// TIA Portal project "latest plc" (V21)

(* hardware
DEVICE "S7-1200 station_1"  S7-1200 Station
   slot 0: "Rack_0"  S7-1200 Rack  Rack  V1.0
   slot 1: "PLC_1"  CPU 1214C DC/DC/DC  6ES7 214-1AG40-0XB0  V4.4
DEVICE "HMI_1"  KTP700 Basic PN
   slot 0: "HMI_1"  KTP700 Basic PN  6AV2 123-2GB03-0AX0  17.0.0.0
   slot 1: "HMI_RT_1"  KTP700 Basic PN  6AV2 123-2GB03-0AX0  17.0.0.0
   slot 5: "HMI_1.IE_CP_1"  PROFINET Interface  17.0.0.0
      slot 1: "PROFINET Interface_1"  PROFINET Interface
         slot 1: "Port_1"  Port
*)

// ===== PLC "PLC_1"  CPU 1214C DC/DC/DC =====

VAR_GLOBAL   // PLC tag table "Default tag table"
   "System_Byte" AT %MB1 : Byte;
   "FirstScan" AT %M1.0 : Bool;
   "DiagStatusUpdate" AT %M1.1 : Bool;
   "AlwaysTRUE" AT %M1.2 : Bool;
   "AlwaysFALSE" AT %M1.3 : Bool;
   "Clock_Byte" AT %MB0 : Byte;
   "Clock_10Hz" AT %M0.0 : Bool;
   "Clock_5Hz" AT %M0.1 : Bool;
   "Clock_2.5Hz" AT %M0.2 : Bool;
   "Clock_2Hz" AT %M0.3 : Bool;
   "Clock_1.25Hz" AT %M0.4 : Bool;
   "Clock_1Hz" AT %M0.5 : Bool;
   "Clock_0.625Hz" AT %M0.6 : Bool;
   "Clock_0.5Hz" AT %M0.7 : Bool;
   "CONTROL ON FLAG" AT %M2.0 : Bool;
   "MANUAL MODE SELECTED" AT %M2.1 : Bool;
   "AUTO MODE SELECTED" AT %M2.2 : Bool;
   "FAULT RESET FLAG" AT %M2.3 : Bool;
   "FAULT BIT" AT %M2.4 : Bool;
   "MANUAL CONVEYOR FWD ON FLAG" AT %M2.5 : Bool;
   "MANUAL CONVEYOR REV ON FLAG" AT %M2.6 : Bool;
END_VAR

VAR_GLOBAL   // PLC tag table "DI"
   "DI_PRODUCT SENSOR" AT %I0.0 : Bool;
   "DI_AUTO MANUAL SELECTION" AT %I0.1 : Bool;
   "DI_CYCLE START PB" AT %I0.2 : Bool;
   "DI_CYCLE STOP PB" AT %I0.3 : Bool;
   "DI_EMERGENCY PB" AT %I0.4 : Bool;
   "DI_CONVEYOR VFD FAULT" AT %I0.5 : Bool;
   "DI_SPARE I0.6" AT %I0.6 : Bool;
   "DI_SPARE I0.7" AT %I0.7 : Bool;
   "DI_SPARE I1.0" AT %I1.0 : Bool;
   "DI_SPARE I1.1" AT %I1.1 : Bool;
   "DI_SPARE I1.2" AT %I1.2 : Bool;
   "DI_SPARE I1.3" AT %I1.3 : Bool;
   "DI_SPARE I1.4" AT %I1.4 : Bool;
   "DI_SPARE I1.5" AT %I1.5 : Bool;
END_VAR

VAR_GLOBAL   // PLC tag table "DO"
   "DO_CONVEYOR FWD ON" AT %Q0.0 : Bool;
   "DO_CONVEYOR REV ON" AT %Q0.1 : Bool;
   "DO_FAULT RESET" AT %Q0.2 : Bool;
   "DO_TL GREEN" AT %Q0.3 : Bool;
   "DO_TL RED" AT %Q0.4 : Bool;
   "DO_TL AMBER" AT %Q0.5 : Bool;
   "DO_SPARE Q0.6" AT %Q0.6 : Bool;
   "DO_SPARE Q0.7" AT %Q0.7 : Bool;
   "DO_SPARE Q1.0" AT %Q1.0 : Bool;
   "DO_SPARE Q1.1" AT %Q1.1 : Bool;
END_VAR

DATA_BLOCK "DB_HMI"   // DB1
{ S7_Optimized_Access := 'FALSE' }
VERSION : 0.1
   VAR
      "FAULT RESET PB" : Bool;
      "MOTOR JOG FWD PB" : Bool;
      "MOTOR JOG REV PB" : Bool;
      "STOP TIME" : DInt;
      "CAMERA DONE" : Bool;
   END_VAR
BEGIN
END_DATA_BLOCK

DATA_BLOCK "DB_ALARMS"   // DB2
{ S7_Optimized_Access := 'FALSE' }
VERSION : 0.1
   VAR
      "EMERGENCY PB PRESSED FAULT" : Bool;
      "VFD FAULT" : Bool;
      SPARE1 : Bool;
      SPARE2 : Bool;
      SPARE3 : Bool;
      SPARE4 : Bool;
      SPARE5 : Bool;
      SPARE6 : Bool;
      SPARE7 : Bool;
      SPARE8 : Bool;
      SPARE9 : Bool;
      SPARE10 : Bool;
      SPARE11 : Bool;
      SPARE12 : Bool;
      SPARE13 : Bool;
      SPARE14 : Bool;
      "FAULT POP" : Bool;
      "WARNING POP" : Bool;
   END_VAR
BEGIN
END_DATA_BLOCK

DATA_BLOCK "DB_AUTO"   // DB3
{ S7_Optimized_Access := 'FALSE' }
VERSION : 0.1
   VAR
      ACTIVE : Bool;
      "CONVEYOR ON" : Bool;
      "CONVEYOR OFF1" : Bool;
      "CONVEYOR OFF2" : Bool;
      P_TRG : Bool;
      "CAMERA DONE" : Bool;
      "AUTO STATUS" : Int;
      "STOP DELAY TIMER" : IEC_TIMER;
      "SENSOR CHECK DELAY" : IEC_TIMER;
   END_VAR
BEGIN
END_DATA_BLOCK

DATA_BLOCK "DB_CAMERA"   // DB5
{ S7_Optimized_Access := 'FALSE' }
VERSION : 0.1
   VAR
      DATA1 : Int;
      DATA2 : Int;
      DATA3 : Int;
      DATA4 : Int;
      DATA5 : Int;
      DATA6 : Int;
      DATA7 : Int;
      DATA8 : Int;
      DATA9 : Int;
      DATA10 : Int;
      DATA11 : Int;
      DATA12 : Int;
      DATA13 : Int;
      DATA14 : Int;
      DATA15 : Int;
      DATA16 : Int;
      DATA17 : Int;
      DATA18 : Int;
      DATA19 : Int;
   END_VAR
BEGIN
END_DATA_BLOCK

DATA_BLOCK "DB_TCP_IP"   // DB12
{ S7_Optimized_Access := 'TRUE' }
VERSION : 0.1
   VAR
      "MY CONNECT DATA" : TCON_IP_v4;
      "NO OF DONE" : UDInt;
      "NO OF ERROR" : UDInt;
      "ERROR STATUS" : UDInt;
   END_VAR
BEGIN
END_DATA_BLOCK

FUNCTION "FC_GENERAL" : Void   // FC1, LAD
{ S7_Optimized_Access := 'TRUE' }
VERSION : 0.1
BEGIN

REGION Network 1: CONTROL ON
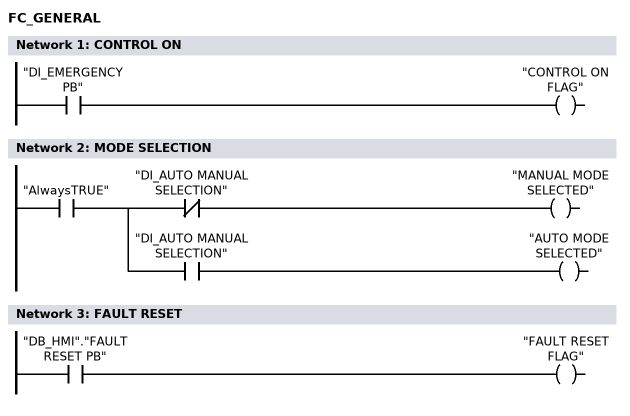
   RUNG wire#powerrail
      Contact( "DI_EMERGENCY PB" )
      Coil( "CONTROL ON FLAG" )
   END_RUNG
   // the same network as SCL:
   "CONTROL ON FLAG" := "DI_EMERGENCY PB";
END_REGION

REGION Network 2: MODE SELECTION
   RUNG wire#powerrail
      Contact( "AlwaysTRUE" )
      wire#w1
      I_Contact( "DI_AUTO MANUAL SELECTION" )
      Coil( "MANUAL MODE SELECTED" )
   END_RUNG
   RUNG wire#w1
      Contact( "DI_AUTO MANUAL SELECTION" )
      Coil( "AUTO MODE SELECTED" )
   END_RUNG
   // the same network as SCL:
   "MANUAL MODE SELECTED" := "AlwaysTRUE" AND NOT "DI_AUTO MANUAL SELECTION";
   "AUTO MODE SELECTED" := "AlwaysTRUE" AND "DI_AUTO MANUAL SELECTION";
END_REGION

REGION Network 3: FAULT RESET
   RUNG wire#powerrail
      Contact( "DB_HMI"."FAULT RESET PB" )
      Coil( "FAULT RESET FLAG" )
   END_RUNG
   // the same network as SCL:
   "FAULT RESET FLAG" := "DB_HMI"."FAULT RESET PB";
END_REGION
END_FUNCTION

FUNCTION "FC_MANUAL" : Void   // FC2, LAD
{ S7_Optimized_Access := 'TRUE' }
VERSION : 0.1
   VAR_TEMP   // added for the SCL form of the ladder/FBD networks
      _w1 : Bool;
   END_VAR
BEGIN

REGION Network 1: MOTOR FWD /REV ON
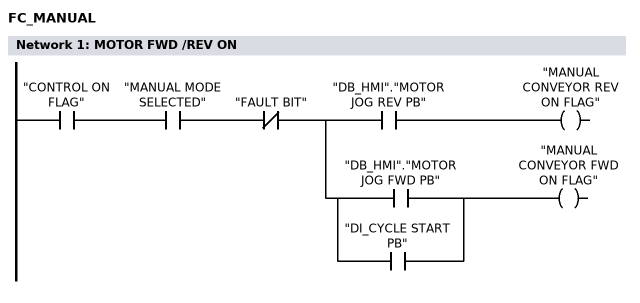
   RUNG wire#powerrail
      Contact( "CONTROL ON FLAG" )
      Contact( "MANUAL MODE SELECTED" )
      I_Contact( "FAULT BIT" )
      wire#w1
      Contact( "DB_HMI"."MOTOR JOG REV PB" )
      Coil( "MANUAL CONVEYOR REV ON FLAG" )
   END_RUNG
   RUNG wire#w1
      Contact( "DB_HMI"."MOTOR JOG FWD PB" )
      wire#w2
      Coil( "MANUAL CONVEYOR FWD ON FLAG" )
   END_RUNG
   RUNG wire#w1
      Contact( "DI_CYCLE START PB" )
   END_RUNG wire#w2
   // the same network as SCL:
   #_w1 := "CONTROL ON FLAG" AND "MANUAL MODE SELECTED" AND NOT "FAULT BIT";
   "MANUAL CONVEYOR REV ON FLAG" := #_w1 AND "DB_HMI"."MOTOR JOG REV PB";
   "MANUAL CONVEYOR FWD ON FLAG" := #_w1 AND ("DB_HMI"."MOTOR JOG FWD PB" OR "DI_CYCLE START PB");
END_REGION
END_FUNCTION

FUNCTION "FC_ALARMS" : Void   // FC3, LAD
{ S7_Optimized_Access := 'TRUE' }
VERSION : 0.1
BEGIN

REGION Network 1: EMERGENCY PB PRESSED FAULT (I0.4)
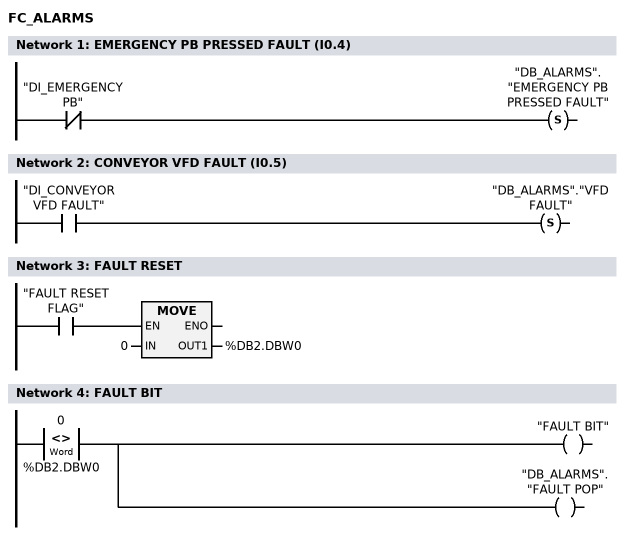
   RUNG wire#powerrail
      I_Contact( "DI_EMERGENCY PB" )
      S_Coil( "DB_ALARMS"."EMERGENCY PB PRESSED FAULT" )
   END_RUNG
   // the same network as SCL:
   IF NOT "DI_EMERGENCY PB" THEN "DB_ALARMS"."EMERGENCY PB PRESSED FAULT" := TRUE; END_IF;
END_REGION

REGION Network 2: CONVEYOR VFD FAULT (I0.5)
   RUNG wire#powerrail
      Contact( "DI_CONVEYOR VFD FAULT" )
      S_Coil( "DB_ALARMS"."VFD FAULT" )
   END_RUNG
   // the same network as SCL:
   IF "DI_CONVEYOR VFD FAULT" THEN "DB_ALARMS"."VFD FAULT" := TRUE; END_IF;
END_REGION

REGION Network 3: FAULT RESET
   RUNG wire#powerrail
      Contact( "FAULT RESET FLAG" )
      Move(in := 0, out1 => %DB2.DBW0)
   END_RUNG
   // the same network as SCL:
   IF "FAULT RESET FLAG" THEN %DB2.DBW0 := 0; END_IF;
END_REGION

REGION Network 4: FAULT BIT
   RUNG wire#powerrail
      { S7_Templates := "SrcType := Word" } NE_Contact(in1 := 0, in2 := %DB2.DBW0)
      wire#w1
      Coil( "FAULT BIT" )
   END_RUNG
   RUNG wire#w1
      Coil( "DB_ALARMS"."FAULT POP" )
   END_RUNG
   // the same network as SCL:
   "FAULT BIT" := 0 <> %DB2.DBW0;
   "DB_ALARMS"."FAULT POP" := "FAULT BIT";
END_REGION
END_FUNCTION

FUNCTION "FC_OUTPUTS" : Void   // FC4, LAD
{ S7_Optimized_Access := 'TRUE' }
VERSION : 0.1
BEGIN

REGION Network 1: CONVEYOR FWD ON
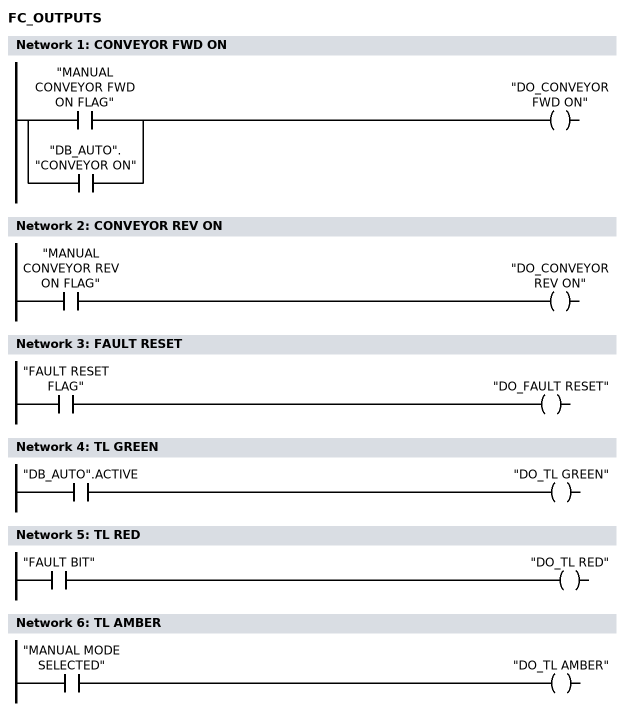
   RUNG wire#powerrail
      Contact( "MANUAL CONVEYOR FWD ON FLAG" )
      wire#w1
      Coil( "DO_CONVEYOR FWD ON" )
   END_RUNG
   RUNG wire#powerrail
      Contact( "DB_AUTO"."CONVEYOR ON" )
   END_RUNG wire#w1
   // the same network as SCL:
   "DO_CONVEYOR FWD ON" := "MANUAL CONVEYOR FWD ON FLAG" OR "DB_AUTO"."CONVEYOR ON";
END_REGION

REGION Network 2: CONVEYOR REV ON
   RUNG wire#powerrail
      Contact( "MANUAL CONVEYOR REV ON FLAG" )
      Coil( "DO_CONVEYOR REV ON" )
   END_RUNG
   // the same network as SCL:
   "DO_CONVEYOR REV ON" := "MANUAL CONVEYOR REV ON FLAG";
END_REGION

REGION Network 3: FAULT RESET
   RUNG wire#powerrail
      Contact( "FAULT RESET FLAG" )
      Coil( "DO_FAULT RESET" )
   END_RUNG
   // the same network as SCL:
   "DO_FAULT RESET" := "FAULT RESET FLAG";
END_REGION

REGION Network 4: TL GREEN
   RUNG wire#powerrail
      Contact( "DB_AUTO".ACTIVE )
      Coil( "DO_TL GREEN" )
   END_RUNG
   // the same network as SCL:
   "DO_TL GREEN" := "DB_AUTO".ACTIVE;
END_REGION

REGION Network 5: TL RED
   RUNG wire#powerrail
      Contact( "FAULT BIT" )
      Coil( "DO_TL RED" )
   END_RUNG
   // the same network as SCL:
   "DO_TL RED" := "FAULT BIT";
END_REGION

REGION Network 6: TL AMBER
   RUNG wire#powerrail
      Contact( "MANUAL MODE SELECTED" )
      Coil( "DO_TL AMBER" )
   END_RUNG
   // the same network as SCL:
   "DO_TL AMBER" := "MANUAL MODE SELECTED";
END_REGION
END_FUNCTION

FUNCTION "FC_AUTO" : Void   // FC5, LAD
{ S7_Optimized_Access := 'TRUE' }
VERSION : 0.1
   VAR_TEMP   // added for the SCL form of the ladder/FBD networks
      _w1 : Bool;
      _w2 : Bool;
      _w3 : Bool;
   END_VAR
BEGIN

REGION Network 1: AUTO ON
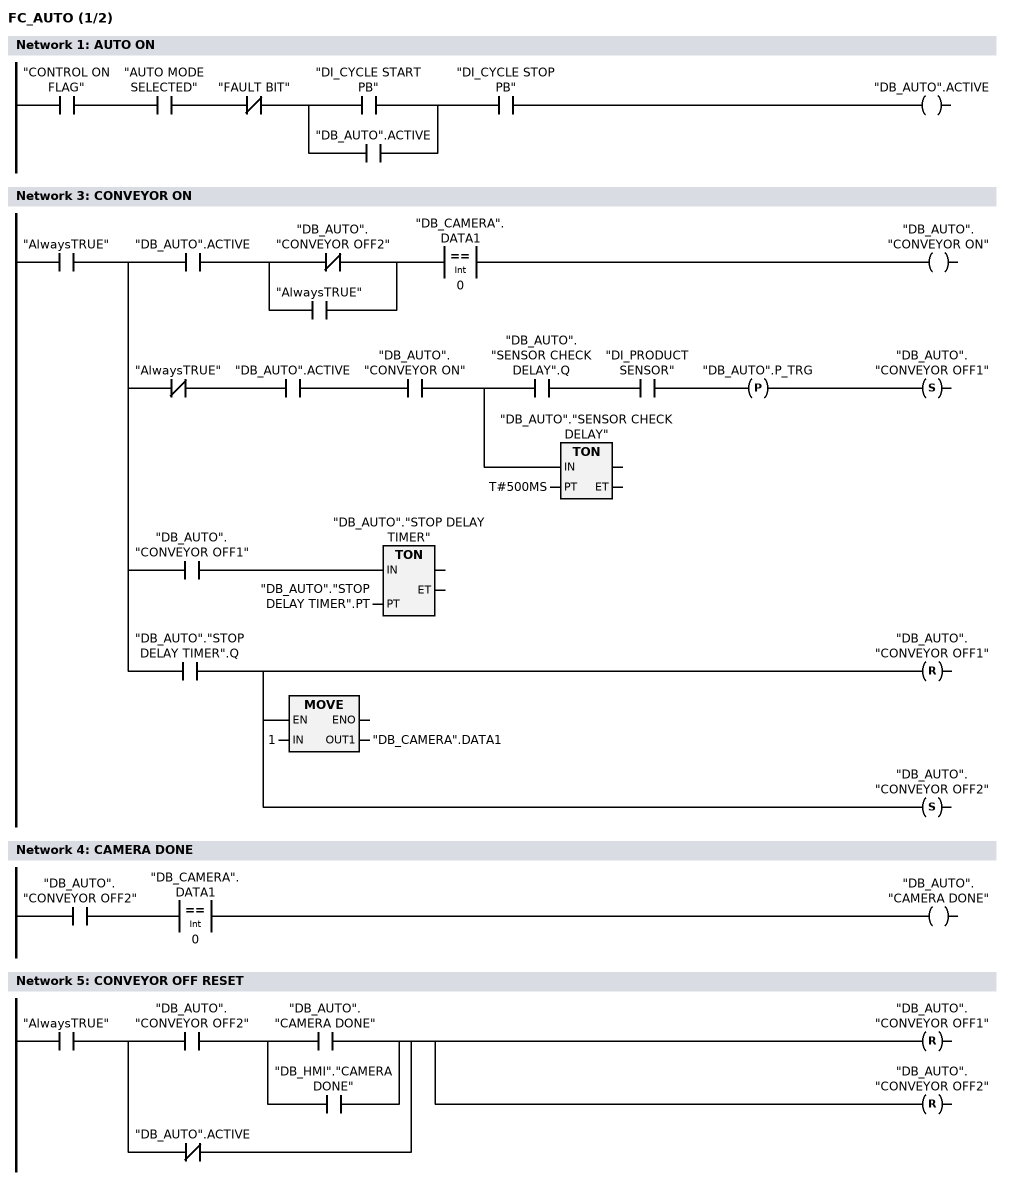
   RUNG wire#powerrail
      Contact( "CONTROL ON FLAG" )
      Contact( "AUTO MODE SELECTED" )
      I_Contact( "FAULT BIT" )
      wire#w1
      Contact( "DI_CYCLE START PB" )
      wire#w2
      Contact( "DI_CYCLE STOP PB" )
      Coil( "DB_AUTO".ACTIVE )
   END_RUNG
   RUNG wire#w1
      Contact( "DB_AUTO".ACTIVE )
   END_RUNG wire#w2
   // the same network as SCL:
   "DB_AUTO".ACTIVE := "CONTROL ON FLAG" AND "AUTO MODE SELECTED" AND NOT "FAULT BIT" AND ("DI_CYCLE START PB" OR "DB_AUTO".ACTIVE) AND "DI_CYCLE STOP PB";
END_REGION

REGION Network 2 (SCL): STOP DELAY TIME
   "DB_AUTO"."STOP DELAY TIMER".PT := "DB_HMI"."STOP TIME" * 1000;
END_REGION

REGION Network 3: CONVEYOR ON
   "DB_AUTO"."CONVEYOR ON" := "AlwaysTRUE" AND "DB_AUTO".ACTIVE AND (NOT "DB_AUTO"."CONVEYOR OFF2" OR "AlwaysTRUE") AND ("DB_CAMERA".DATA1 = 0);
   #_w1 := "AlwaysTRUE" AND NOT "AlwaysTRUE" AND "DB_AUTO".ACTIVE AND "DB_AUTO"."CONVEYOR ON";
   #_w2 := #_w1 AND "DB_AUTO"."SENSOR CHECK DELAY".Q AND "DI_PRODUCT SENSOR";
   #_w3 := #_w2 AND NOT "DB_AUTO".P_TRG;   // rising edge
   "DB_AUTO".P_TRG := #_w2;
   IF #_w3 THEN "DB_AUTO"."CONVEYOR OFF1" := TRUE; END_IF;
   "DB_AUTO"."SENSOR CHECK DELAY".TON(IN := #_w1, PT := T#500MS);
   "DB_AUTO"."STOP DELAY TIMER".TON(IN := "AlwaysTRUE" AND "DB_AUTO"."CONVEYOR OFF1",
                           PT := "DB_AUTO"."STOP DELAY TIMER".PT);
   IF "AlwaysTRUE" AND "DB_AUTO"."STOP DELAY TIMER".Q THEN
       "DB_AUTO"."CONVEYOR OFF1" := FALSE;
       "DB_CAMERA".DATA1 := 1;
       "DB_AUTO"."CONVEYOR OFF2" := TRUE;
   END_IF;
END_REGION

REGION Network 4: CAMERA DONE
   RUNG wire#powerrail
      Contact( "DB_AUTO"."CONVEYOR OFF2" )
      { S7_Templates := "SrcType := Int" } EQ_Contact(in1 := "DB_CAMERA".DATA1, in2 := 0)
      Coil( "DB_AUTO"."CAMERA DONE" )
   END_RUNG
   // the same network as SCL:
   "DB_AUTO"."CAMERA DONE" := "DB_AUTO"."CONVEYOR OFF2" AND ("DB_CAMERA".DATA1 = 0);
END_REGION

REGION Network 5: CONVEYOR OFF RESET
   RUNG wire#powerrail
      Contact( "AlwaysTRUE" )
      wire#w1
      Contact( "DB_AUTO"."CONVEYOR OFF2" )
      wire#w2
      Contact( "DB_AUTO"."CAMERA DONE" )
      wire#w3
      R_Coil( "DB_AUTO"."CONVEYOR OFF1" )
   END_RUNG
   RUNG wire#w2
      Contact( "DB_HMI"."CAMERA DONE" )
   END_RUNG wire#w3
   RUNG wire#w1
      I_Contact( "DB_AUTO".ACTIVE )
   END_RUNG wire#w3
   RUNG wire#w3
      R_Coil( "DB_AUTO"."CONVEYOR OFF2" )
   END_RUNG
   // the same network as SCL:
   IF "AlwaysTRUE" AND (("DB_AUTO"."CONVEYOR OFF2" AND ("DB_AUTO"."CAMERA DONE" OR "DB_HMI"."CAMERA DONE")) OR NOT "DB_AUTO".ACTIVE) THEN
       "DB_AUTO"."CONVEYOR OFF1" := FALSE;
       "DB_AUTO"."CONVEYOR OFF2" := FALSE;
   END_IF;
END_REGION

REGION Network 6: AUTO STATUS
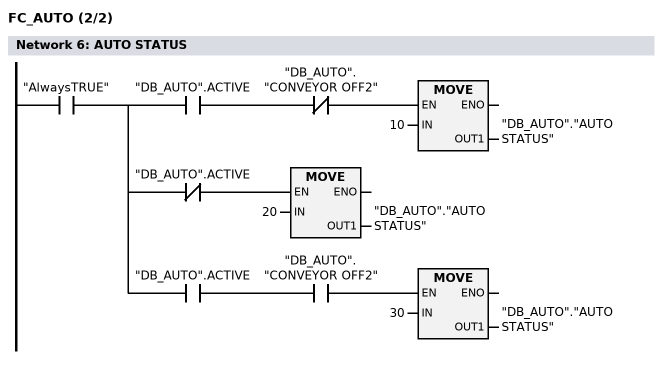
   RUNG wire#powerrail
      Contact( "AlwaysTRUE" )
      wire#w1
      Contact( "DB_AUTO".ACTIVE )
      I_Contact( "DB_AUTO"."CONVEYOR OFF2" )
      Move(in := 10, out1 => "DB_AUTO"."AUTO STATUS")
   END_RUNG
   RUNG wire#w1
      I_Contact( "DB_AUTO".ACTIVE )
      Move(in := 20, out1 => "DB_AUTO"."AUTO STATUS")
   END_RUNG
   RUNG wire#w1
      Contact( "DB_AUTO".ACTIVE )
      Contact( "DB_AUTO"."CONVEYOR OFF2" )
      Move(in := 30, out1 => "DB_AUTO"."AUTO STATUS")
   END_RUNG
   // the same network as SCL:
   IF "AlwaysTRUE" AND "DB_AUTO".ACTIVE AND NOT "DB_AUTO"."CONVEYOR OFF2" THEN
       "DB_AUTO"."AUTO STATUS" := 10;
   END_IF;
   IF "AlwaysTRUE" AND NOT "DB_AUTO".ACTIVE THEN "DB_AUTO"."AUTO STATUS" := 20; END_IF;
   IF "AlwaysTRUE" AND "DB_AUTO".ACTIVE AND "DB_AUTO"."CONVEYOR OFF2" THEN
       "DB_AUTO"."AUTO STATUS" := 30;
   END_IF;
END_REGION
END_FUNCTION

FUNCTION "FC_TCP_IP" : Void   // FC6, LAD
{ S7_Optimized_Access := 'TRUE' }
VERSION : 0.1
BEGIN

REGION Network 1: Connection definition
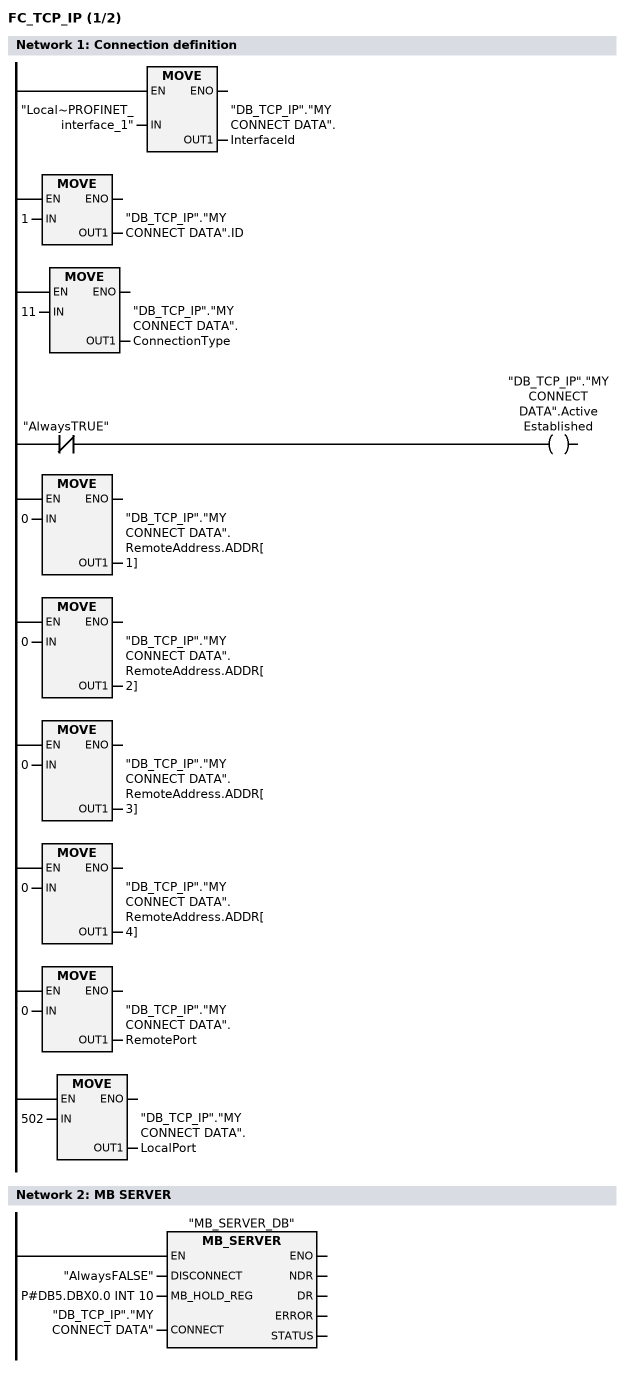
   RUNG wire#powerrail
      Move(in := "Local~PROFINET_interface_1", out1 => "DB_TCP_IP"."MY CONNECT DATA".InterfaceId)
   END_RUNG
   RUNG wire#powerrail
      Move(in := 1, out1 => "DB_TCP_IP"."MY CONNECT DATA".ID)
   END_RUNG
   RUNG wire#powerrail
      Move(in := 11, out1 => "DB_TCP_IP"."MY CONNECT DATA".ConnectionType)
   END_RUNG
   RUNG wire#powerrail
      I_Contact( "AlwaysTRUE" )
      Coil( "DB_TCP_IP"."MY CONNECT DATA".ActiveEstablished )
   END_RUNG
   RUNG wire#powerrail
      Move(in := 0, out1 => "DB_TCP_IP"."MY CONNECT DATA".RemoteAddress.ADDR[1])
   END_RUNG
   RUNG wire#powerrail
      Move(in := 0, out1 => "DB_TCP_IP"."MY CONNECT DATA".RemoteAddress.ADDR[2])
   END_RUNG
   RUNG wire#powerrail
      Move(in := 0, out1 => "DB_TCP_IP"."MY CONNECT DATA".RemoteAddress.ADDR[3])
   END_RUNG
   RUNG wire#powerrail
      Move(in := 0, out1 => "DB_TCP_IP"."MY CONNECT DATA".RemoteAddress.ADDR[4])
   END_RUNG
   RUNG wire#powerrail
      Move(in := 0, out1 => "DB_TCP_IP"."MY CONNECT DATA".RemotePort)
   END_RUNG
   RUNG wire#powerrail
      Move(in := 502, out1 => "DB_TCP_IP"."MY CONNECT DATA".LocalPort)
   END_RUNG
   // the same network as SCL:
   "DB_TCP_IP"."MY CONNECT DATA".InterfaceId := "Local~PROFINET_interface_1";
   "DB_TCP_IP"."MY CONNECT DATA".ID := 1;
   "DB_TCP_IP"."MY CONNECT DATA".ConnectionType := 11;
   "DB_TCP_IP"."MY CONNECT DATA".ActiveEstablished := NOT "AlwaysTRUE";
   "DB_TCP_IP"."MY CONNECT DATA".RemoteAddress.ADDR[1] := 0;
   "DB_TCP_IP"."MY CONNECT DATA".RemoteAddress.ADDR[2] := 0;
   "DB_TCP_IP"."MY CONNECT DATA".RemoteAddress.ADDR[3] := 0;
   "DB_TCP_IP"."MY CONNECT DATA".RemoteAddress.ADDR[4] := 0;
   "DB_TCP_IP"."MY CONNECT DATA".RemotePort := 0;
   "DB_TCP_IP"."MY CONNECT DATA".LocalPort := 502;
END_REGION

REGION Network 2: MB SERVER
   "MB_SERVER_DB"(DISCONNECT := "AlwaysFALSE",   // MB_SERVER
                  MB_HOLD_REG := P#DB5.DBX0.0 INT 10,
                  CONNECT := "DB_TCP_IP"."MY CONNECT DATA");
END_REGION

REGION Network 3: ERROR CHECK
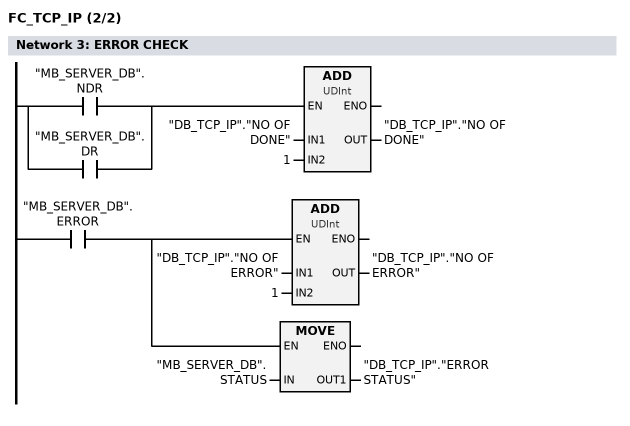
   RUNG wire#powerrail
      Contact( "MB_SERVER_DB".NDR )
      wire#w1
      { S7_Templates := "SrcType := UDInt" } Add(in1 := "DB_TCP_IP"."NO OF DONE", in2 := 1, out => "DB_TCP_IP"."NO OF DONE")
   END_RUNG
   RUNG wire#powerrail
      Contact( "MB_SERVER_DB".DR )
   END_RUNG wire#w1
   RUNG wire#powerrail
      Contact( "MB_SERVER_DB".ERROR )
      wire#w2
      { S7_Templates := "SrcType := UDInt" } Add(in1 := "DB_TCP_IP"."NO OF ERROR", in2 := 1, out => "DB_TCP_IP"."NO OF ERROR")
   END_RUNG
   RUNG wire#w2
      Move(in := "MB_SERVER_DB".STATUS, out1 => "DB_TCP_IP"."ERROR STATUS")
   END_RUNG
   // the same network as SCL:
   IF "MB_SERVER_DB".NDR OR "MB_SERVER_DB".DR THEN
       "DB_TCP_IP"."NO OF DONE" := "DB_TCP_IP"."NO OF DONE" + 1;
   END_IF;
   IF "MB_SERVER_DB".ERROR THEN
       "DB_TCP_IP"."NO OF ERROR" := "DB_TCP_IP"."NO OF ERROR" + 1;
       "DB_TCP_IP"."ERROR STATUS" := "MB_SERVER_DB".STATUS;
   END_IF;
END_REGION
END_FUNCTION

ORGANIZATION_BLOCK "Main"   // OB1, LAD, ProgramCycle
TITLE = "Main Program Sweep (Cycle)"
{ S7_Optimized_Access := 'TRUE' }
VERSION : 0.1
   VAR_INPUT
      Initial_Call : Bool;   // Initial call of this OB
      Remanence : Bool;   // =True, if remanent data are available
   END_VAR
BEGIN

REGION Network 1
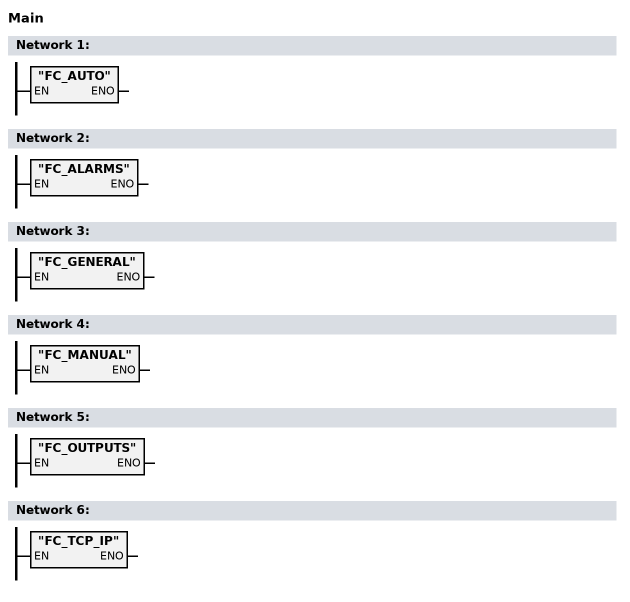
   RUNG wire#powerrail
      "FC_AUTO"()
   END_RUNG
   // the same network as SCL:
   "FC_AUTO"();
END_REGION

REGION Network 2
   RUNG wire#powerrail
      "FC_ALARMS"()
   END_RUNG
   // the same network as SCL:
   "FC_ALARMS"();
END_REGION

REGION Network 3
   RUNG wire#powerrail
      "FC_GENERAL"()
   END_RUNG
   // the same network as SCL:
   "FC_GENERAL"();
END_REGION

REGION Network 4
   RUNG wire#powerrail
      "FC_MANUAL"()
   END_RUNG
   // the same network as SCL:
   "FC_MANUAL"();
END_REGION

REGION Network 5
   RUNG wire#powerrail
      "FC_OUTPUTS"()
   END_RUNG
   // the same network as SCL:
   "FC_OUTPUTS"();
END_REGION

REGION Network 6
   RUNG wire#powerrail
      "FC_TCP_IP"()
   END_RUNG
   // the same network as SCL:
   "FC_TCP_IP"();
END_REGION
END_ORGANIZATION_BLOCK

(* ===== HMI "HMI_RT_1" =====
system functions are stored by id; their names below are inferred from use
connection "HMI_Connection_1": ETHERNET, SMART_S7_1200_OMS

HMI tags "Default tag table"
   "Tag_ScreenNumber" : UInt, internal
   "AUTO MODE SELECTED" : Bool = PLC "AUTO MODE SELECTED" AT %M2.2, 1 s
   "DB_ALARMS_FAULT POP" : Bool = PLC DB_ALARMS."FAULT POP" AT %DB2.DBX2.0, 1 s
   "DB_ALARMS_WARNING POP" : Bool = PLC DB_ALARMS."WARNING POP" AT %DB2.DBX2.1, 1 s
   "DB_HMI_FAULT RESET PB" : Bool = PLC DB_HMI."FAULT RESET PB" AT %DB1.DBX0.0, 1 s
   "DB_HMI_MOTOR JOG FWD PB" : Bool = PLC DB_HMI."MOTOR JOG FWD PB" AT %DB1.DBX0.1, 1 s
   "DB_HMI_MOTOR JOG REV PB" : Bool = PLC DB_HMI."MOTOR JOG REV PB" AT %DB1.DBX0.2, 1 s
   "DB_AUTO_AUTO STATUS" : Int = PLC DB_AUTO."AUTO STATUS" AT %DB3.DBW2, 1 s
   "DB_HMI_STOP TIME" : DInt = PLC DB_HMI."STOP TIME" AT %DB1.DBD2, 1 s
   "DB_HMI_CAMERA DONE" : Bool = PLC DB_HMI."CAMERA DONE" AT %DB1.DBX6.0, 1 s

HMI tags "IO"
   "IB0" : Byte AT %IB0, 1 s
   "IB1" : Byte AT %IB1, 1 s
   "QB0" : Byte AT %QB0, 1 s
   "QB1" : Byte AT %QB1, 1 s

HMI tags "ALARMS"
   "ALARM WORD" : Int AT %DB2.DBW0, 1 s

discrete alarms
   1: 'EMERGENCY PB PRESSED FAULT (I0.4)', class Errors, trigger "ALARM WORD" bit 8
   2: 'CONVEYOR VFD FAULT (I0.5)', class Errors, trigger "ALARM WORD" bit 9
   3: '', class Errors, trigger "ALARM WORD" bit 10
   4: '', class Errors, trigger "ALARM WORD" bit 11
   5: '', class Errors, trigger "ALARM WORD" bit 12
   6: '', class Errors, trigger "ALARM WORD" bit 13
   7: '', class Errors, trigger "ALARM WORD" bit 14
   8: '', class Errors, trigger "ALARM WORD" bit 15

text list "AUTO STATUS": 10 'AUTO RUNNING'; 20 'STOPPED'; 30 'WAITING FOR CAMERA ACK'

text list "MODE": 0 'MANUAL'; 1 'AUTO'

screen "AUTO" 800x480, template "MAIN"
   TextField "Template_Text field_2" at 308,62 size 181x27; Text 'AUTO OPERATION'
   SymbolicIOField "Symbolic I/O field_1" at 116,182 size 560x106; TextOff '0'; TextOn '1'; TextList "AUTO STATUS"
      ProcessValue <- "DB_AUTO_AUTO STATUS"
      Appearance <- "DB_AUTO_AUTO STATUS"
   TextField "Template_Text field_1" at 304,117 size 165x34; Text 'AUTO STATUS'

Template "MAIN" 800x480
   DateTimeField "HmiScreenItemData" at 1,1 size 121x58
   DateTimeField "HmiScreenItemData_1" at 677,1 size 121x58
   Button "Template_Button_1" at 6,411 size 151x60; TextOff 'AUTO'
      on Press: ActivateScreen("AUTO", 0)
   Button "Template_Button_7" at 0,61 size 800x30; TextOff 'Text'
   TextField "Template_Text field_1" at 225,11 size 327x39; Text 'CONVEYOR'
   TextField "Template_Text field_2" at 12,64 size 65x23; Text 'MODE :-'
   SymbolicIOField "Template_Symbolic I/O field_1" at 89,61 size 117x27; TextOff '0'; TextOn '1'; TextList "MODE"
      ProcessValue <- "AUTO MODE SELECTED"
   Button "Template_Button_2" at 166,411 size 151x60; TextOff 'MANUAL'
      on Press: ActivateScreen("MANUAL", 0)
   Button "Template_Button_3" at 326,411 size 151x60; TextOff 'ALARMS'
      on Press: ActivateScreen("ALARMS", 0)
   Button "Template_Button_4" at 486,411 size 151x60; TextOff 'IO STATUS'
      on Press: ActivateScreen("INPUT STATUS", 0)
   Button "Template_Button_5" at 646,411 size 151x60; TextOff 'FAULT RESET'
      on Press: function_b14e0dd5("DB_HMI_FAULT RESET PB", 0)
   AlarmView "Template_Alarm view_2" at 124,4 size 550x53
      Visibility <- "DB_ALARMS_FAULT POP"
   AlarmView "Template_Alarm view_1" at 124,4 size 550x53
      Visibility <- "DB_ALARMS_WARNING POP"

screen "MANUAL" 800x480, template "MAIN"
   Button "Button_1" at 166,194 size 179x82; TextOff 'CONVEYOR FWD JOG'
      on Press: function_b14e0dd5("DB_HMI_MOTOR JOG FWD PB", 0)
      Appearance <- "DB_HMI_MOTOR JOG FWD PB"
   Button "Button_2" at 429,190 size 179x82; TextOff 'CONVEYOR REV JOG'
      Appearance <- "DB_HMI_MOTOR JOG REV PB"
      on Press: function_b14e0dd5("DB_HMI_MOTOR JOG REV PB", 0)
   TextField "Template_Text field_2" at 308,62 size 210x27; Text 'MANUAL OPERATION'

screen "ALARMS" 800x480, template "MAIN"
   AlarmView "Alarm view_1" at 2,92 size 797x308
   TextField "Template_Text field_2" at 372,62 size 84x27; Text 'ALARMS'

screen "INPUT STATUS" 800x480, template "MAIN"
   TextField "Text field_2" at 99,31 size 14x20; Text 'Text'
   TextField "Text field_5" at 0,94 size 84x26; Text 'ADDRESS'
   TextField "Text field_4" at 85,94 size 70x26; Text 'STATUS'
   TextField "Text field_6" at 156,94 size 241x26; Text 'DESCRIPTION'
   TextField "Text field_7" at 156,120 size 242x34; Text 'PRODUCT SENSOR'
   TextField "Text field_8" at 99,31 size 14x20; Text 'Text'
   TextField "Text field_33" at 401,94 size 84x26; Text 'ADDRESS'
   TextField "Text field_34" at 486,94 size 70x26; Text 'STATUS'
   TextField "Text field_35" at 557,94 size 242x26; Text 'DESCRIPTION'
   TextField "Text field_30" at 0,120 size 84x34; Text 'I0.0'
   TextField "Text field_9" at 85,120 size 70x34; Text 'Text'
   TextField "Text field_11" at 156,155 size 242x34; Text 'AUTO MANUAL SELECTION'
   TextField "Text field_12" at 0,155 size 84x34; Text 'I0.1'
   TextField "Text field_13" at 85,155 size 70x34; Text 'Text'
   TextField "Text field_14" at 156,191 size 242x34; Text 'CYCLE START PB'
   TextField "Text field_15" at 0,191 size 84x34; Text 'I0.2'
   TextField "Text field_16" at 85,191 size 70x34; Text 'Text'
   TextField "Text field_17" at 156,227 size 242x34; Text 'CYCLE STOP PB'
   TextField "Text field_18" at 0,227 size 84x34; Text 'I0.3'
   TextField "Text field_19" at 85,227 size 70x34; Text 'Text'
   TextField "Text field_20" at 156,263 size 242x34; Text 'EMERGENCY PB'
   TextField "Text field_21" at 0,263 size 84x34; Text 'I0.4'
   TextField "Text field_22" at 85,263 size 70x34; Text 'Text'
   TextField "Text field_23" at 156,299 size 242x34; Text 'CONVEYOR VFD FAULT'
   TextField "Text field_24" at 0,299 size 84x34; Text 'I0.5'
   TextField "Text field_25" at 85,299 size 70x34; Text 'Text'
   TextField "Text field_26" at 156,335 size 242x34; Text 'SPARE'
   TextField "Text field_27" at 0,335 size 84x34; Text 'I0.6'
   TextField "Text field_28" at 85,335 size 70x34; Text 'Text'
   TextField "Text field_29" at 156,371 size 242x34; Text 'SPARE'
   TextField "Text field_31" at 0,371 size 84x34; Text 'I0.7'
   TextField "Text field_32" at 85,371 size 70x34; Text 'Text'
   TextField "Text field_10" at 557,120 size 242x34; Text 'SPARE'
   TextField "Text field_36" at 401,120 size 84x34; Text 'I1.0'
   TextField "Text field_37" at 486,120 size 70x34; Text 'Text'
   TextField "Text field_38" at 557,155 size 242x34; Text 'SPARE'
   TextField "Text field_39" at 401,155 size 84x34; Text 'I1.1'
   TextField "Text field_40" at 486,155 size 70x34; Text 'Text'
   TextField "Text field_41" at 557,191 size 242x34; Text 'SPARE'
   TextField "Text field_42" at 401,191 size 84x34; Text 'I1.2'
   TextField "Text field_43" at 486,191 size 70x34; Text 'Text'
   TextField "Text field_44" at 557,227 size 242x34; Text 'SPARE'
   TextField "Text field_45" at 401,227 size 84x34; Text 'I1.3'
   TextField "Text field_46" at 486,227 size 70x34; Text 'Text'
   Circle "Circle_1" at 109,126 size 23x23
      Appearance <- "IB0"
   Circle "Circle_2" at 109,161 size 23x23
      Appearance <- "IB0"
   Circle "Circle_3" at 109,197 size 23x23
      Appearance <- "IB0"
   Circle "Circle_4" at 109,233 size 23x23
      Appearance <- "IB0"
   Circle "Circle_5" at 109,269 size 23x23
      Appearance <- "IB0"
   Circle "Circle_6" at 109,305 size 23x23
      Appearance <- "IB0"
   Circle "Circle_7" at 109,341 size 23x23
      Appearance <- "IB0"
   Circle "Circle_8" at 109,377 size 23x23
      Appearance <- "IB0"
   Circle "Circle_9" at 510,126 size 23x23
      Appearance <- "IB1"
   Circle "Circle_10" at 510,161 size 23x23
      Appearance <- "IB1"
   Circle "Circle_11" at 510,197 size 23x23
      Appearance <- "IB1"
   Circle "Circle_12" at 510,233 size 23x23
      Appearance <- "IB1"
   TextField "Text field_3" at 558,263 size 242x34; Text 'SPARE'
   TextField "Text field_47" at 402,263 size 84x34; Text 'I1.4'
   TextField "Text field_48" at 487,263 size 70x34; Text 'Text'
   Circle "Circle_13" at 511,269 size 23x23
      Appearance <- "IB1"
   TextField "Text field_49" at 558,299 size 242x34; Text 'SPARE'
   TextField "Text field_50" at 402,299 size 84x34; Text 'I1.5'
   TextField "Text field_51" at 487,299 size 70x34; Text 'Text'
   Circle "Circle_14" at 511,304 size 23x23
      Appearance <- "IB1"
   TextField "Text field_1" at 308,63 size 147x27; Text 'INPUT STATUS'
   Button "Template_Button_4" at 644,341 size 151x60; TextOff 'NEXT'
      on Press: ActivateScreen("OUTPUT STATUS", 0)

screen "OUTPUT STATUS" 800x480, template "MAIN"
   TextField "Text field_2" at 99,31 size 14x20; Text 'Text'
   TextField "Text field_7" at 156,121 size 242x34; Text 'CONVEYOR FWD ON'
   TextField "Text field_8" at 99,31 size 14x20; Text 'Text'
   TextField "Text field_30" at 0,121 size 84x34; Text 'Q0.0'
   TextField "Text field_9" at 85,121 size 70x34; Text 'Text'
   TextField "Text field_11" at 156,156 size 242x34; Text 'CONVEYOR REV ON'
   TextField "Text field_12" at 0,156 size 84x34; Text 'Q0.1'
   TextField "Text field_13" at 85,156 size 70x34; Text 'Text'
   TextField "Text field_14" at 156,192 size 242x34; Text 'FAULT RESET'
   TextField "Text field_15" at 0,192 size 84x34; Text 'Q0.2'
   TextField "Text field_16" at 85,192 size 70x34; Text 'Text'
   TextField "Text field_17" at 156,228 size 242x34; Text 'TL GREEN'
   TextField "Text field_18" at 0,228 size 84x34; Text 'Q0.3'
   TextField "Text field_19" at 85,228 size 70x34; Text 'Text'
   TextField "Text field_20" at 156,264 size 242x34; Text 'TL RED'
   TextField "Text field_21" at 0,264 size 84x34; Text 'Q0.4'
   TextField "Text field_22" at 85,264 size 70x34; Text 'Text'
   TextField "Text field_23" at 156,300 size 242x34; Text 'TL AMBER'
   TextField "Text field_24" at 0,300 size 84x34; Text 'Q0.5'
   TextField "Text field_25" at 85,300 size 70x34; Text 'Text'
   TextField "Text field_26" at 156,336 size 242x34; Text 'SPARE'
   TextField "Text field_27" at 0,336 size 84x34; Text 'Q0.6'
   TextField "Text field_28" at 85,336 size 70x34; Text 'Text'
   TextField "Text field_29" at 156,372 size 242x34; Text 'SPARE'
   TextField "Text field_31" at 0,372 size 84x34; Text 'Q0.7'
   TextField "Text field_32" at 85,372 size 70x34; Text 'Text'
   TextField "Text field_10" at 557,121 size 242x34; Text 'SPARE'
   TextField "Text field_36" at 401,121 size 84x34; Text 'Q1.0'
   TextField "Text field_37" at 486,121 size 70x34; Text 'Text'
   TextField "Text field_38" at 557,156 size 242x34; Text 'SPARE'
   TextField "Text field_39" at 401,156 size 84x34; Text 'Q1.1'
   TextField "Text field_40" at 486,156 size 70x34; Text 'Text'
   Circle "Circle_1" at 109,127 size 23x23
      Appearance <- "QB0"
   Circle "Circle_2" at 109,162 size 23x23
      Appearance <- "QB0"
   Circle "Circle_3" at 109,198 size 23x23
      Appearance <- "QB0"
   Circle "Circle_4" at 109,234 size 23x23
      Appearance <- "QB0"
   Circle "Circle_5" at 109,270 size 23x23
      Appearance <- "QB0"
   Circle "Circle_6" at 109,306 size 23x23
      Appearance <- "QB0"
   Circle "Circle_7" at 109,342 size 23x23
      Appearance <- "QB0"
   Circle "Circle_8" at 109,378 size 23x23
      Appearance <- "QB0"
   Circle "Circle_9" at 510,127 size 23x23
      Appearance <- "QB1"
   Circle "Circle_10" at 510,162 size 23x23
      Appearance <- "QB1"
   TextField "Text field_1" at 308,63 size 184x27; Text 'OUTPUT STATUS-1'
   TextField "Text field_5" at 0,94 size 84x26; Text 'ADDRESS'
   TextField "Text field_4" at 85,94 size 70x26; Text 'STATUS'
   TextField "Text field_6" at 156,94 size 241x26; Text 'DESCRIPTION'
   TextField "Text field_33" at 401,94 size 84x26; Text 'ADDRESS'
   TextField "Text field_34" at 486,94 size 70x26; Text 'STATUS'
   TextField "Text field_35" at 557,94 size 242x26; Text 'DESCRIPTION'
   Button "Template_Button_4" at 644,341 size 151x60; TextOff 'BACK'
      on Press: ActivateScreen("OUTPUT STATUS", 0)
*)